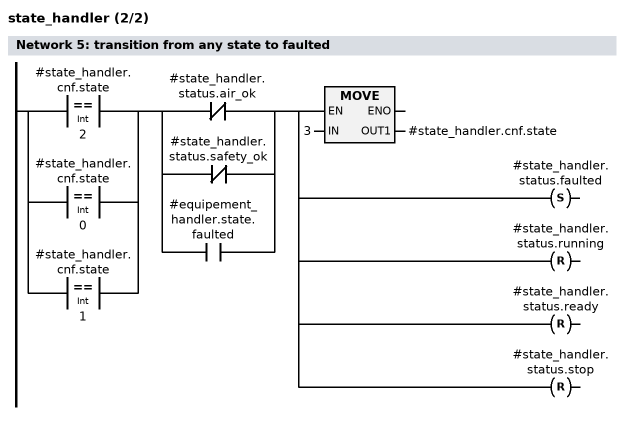
   RUNG wire#powerrail
      { S7_Templates := "SrcType := Int" } EQ_Contact(in1 := #state_handler.cnf.state, in2 := 2)
      wire#w1
      I_Contact( #state_handler.status.air_ok )
      wire#w2
      Move(in := 3, out1 => #state_handler.cnf.state)
   END_RUNG
   RUNG wire#powerrail
      { S7_Templates := "SrcType := Int" } EQ_Contact(in1 := #state_handler.cnf.state, in2 := 0)
   END_RUNG wire#w1
   RUNG wire#powerrail
      { S7_Templates := "SrcType := Int" } EQ_Contact(in1 := #state_handler.cnf.state, in2 := 1)
   END_RUNG wire#w1
   RUNG wire#w1
      I_Contact( #state_handler.status.safety_ok )
   END_RUNG wire#w2
   RUNG wire#w1
      Contact( #equipement_handler.state.faulted )
   END_RUNG wire#w2
   RUNG wire#w2
      S_Coil( #state_handler.status.faulted )
   END_RUNG
   RUNG wire#w2
      R_Coil( #state_handler.status.running )
   END_RUNG
   RUNG wire#w2
      R_Coil( #state_handler.status.ready )
   END_RUNG
   RUNG wire#w2
      R_Coil( #state_handler.status.stop )
   END_RUNG
   // the same network as SCL:
   #_w1 := ((#state_handler.cnf.state = 2) OR (#state_handler.cnf.state = 0) OR (#state_handler.cnf.state = 1)) AND (NOT #state_handler.status.air_ok OR NOT #state_handler.status.safety_ok OR #equipement_handler.state.faulted);
   IF #_w1 THEN
       #state_handler.cnf.state := 3;
       #state_handler.status.faulted := TRUE;
       #state_handler.status.running := FALSE;
       #state_handler.status.ready := FALSE;
       #state_handler.status.stop := FALSE;
   END_IF;
END_REGION
END_FUNCTION_BLOCK

FUNCTION_BLOCK "tower_handler"   // FB3, LAD
{ S7_Optimized_Access := 'TRUE' }
VERSION : 0.1
   VAR_OUTPUT
      tower_green_light : Bool;
      tower_red_light : Bool;
      tower_orange_light : Bool;
      tower_buzer : Bool;
   END_VAR
   VAR_IN_OUT
      state_handler_Machine : "udt_state_handler";
      tower_udt : "udt_tower_handler";
   END_VAR
BEGIN

REGION Network 1: geen light machine is running
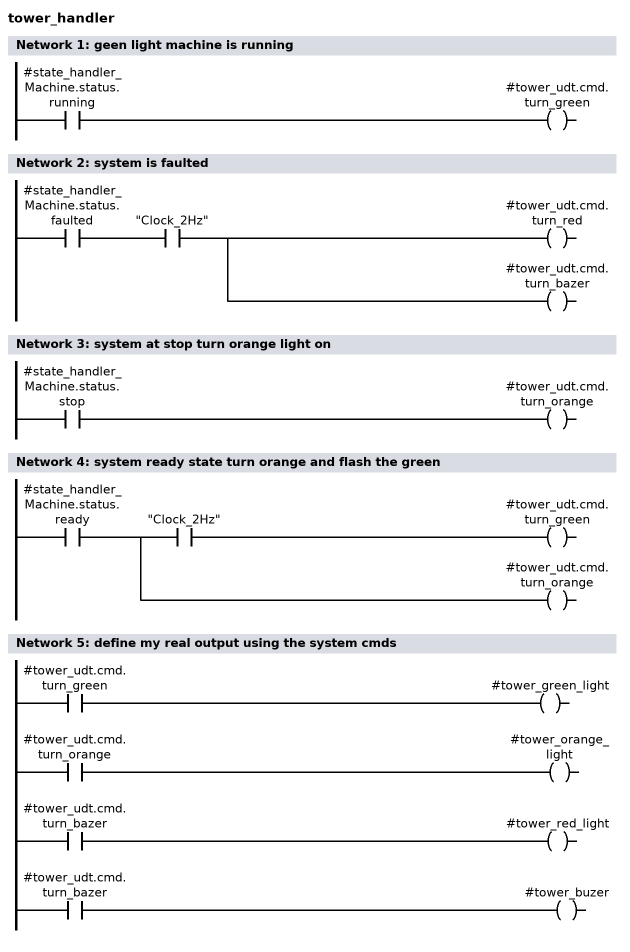
   RUNG wire#powerrail
      Contact( #state_handler_Machine.status.running )
      Coil( #tower_udt.cmd.turn_green )
   END_RUNG
   // the same network as SCL:
   #tower_udt.cmd.turn_green := #state_handler_Machine.status.running;
END_REGION

REGION Network 2: system is faulted
   RUNG wire#powerrail
      Contact( #state_handler_Machine.status.faulted )
      Contact( "Clock_2Hz" )
      wire#w1
      Coil( #tower_udt.cmd.turn_red )
   END_RUNG
   RUNG wire#w1
      Coil( #tower_udt.cmd.turn_bazer )
   END_RUNG
   // the same network as SCL:
   #tower_udt.cmd.turn_red := #state_handler_Machine.status.faulted AND "Clock_2Hz";
   #tower_udt.cmd.turn_bazer := #tower_udt.cmd.turn_red;
END_REGION

REGION Network 3: system at stop turn orange light on
   RUNG wire#powerrail
      Contact( #state_handler_Machine.status.stop )
      Coil( #tower_udt.cmd.turn_orange )
   END_RUNG
   // the same network as SCL:
   #tower_udt.cmd.turn_orange := #state_handler_Machine.status.stop;
END_REGION

REGION Network 4: system ready state turn orange and flash the green
   RUNG wire#powerrail
      Contact( #state_handler_Machine.status.ready )
      wire#w1
      Contact( "Clock_2Hz" )
      Coil( #tower_udt.cmd.turn_green )
   END_RUNG
   RUNG wire#w1
      Coil( #tower_udt.cmd.turn_orange )
   END_RUNG
   // the same network as SCL:
   #tower_udt.cmd.turn_green := #state_handler_Machine.status.ready AND "Clock_2Hz";
   #tower_udt.cmd.turn_orange := #state_handler_Machine.status.ready;
END_REGION

REGION Network 5: define my real output using the system cmds
   RUNG wire#powerrail
      Contact( #tower_udt.cmd.turn_green )
      Coil( #tower_green_light )
   END_RUNG
   RUNG wire#powerrail
      Contact( #tower_udt.cmd.turn_orange )
      Coil( #tower_orange_light )
   END_RUNG
   RUNG wire#powerrail
      Contact( #tower_udt.cmd.turn_bazer )
      Coil( #tower_red_light )
   END_RUNG
   RUNG wire#powerrail
      Contact( #tower_udt.cmd.turn_bazer )
      Coil( #tower_buzer )
   END_RUNG
   // the same network as SCL:
   #tower_green_light := #tower_udt.cmd.turn_green;
   #tower_orange_light := #tower_udt.cmd.turn_orange;
   #tower_red_light := #tower_udt.cmd.turn_bazer;
   #tower_buzer := #tower_udt.cmd.turn_bazer;
END_REGION
END_FUNCTION_BLOCK

FUNCTION_BLOCK "safety_block"   // FB4, LAD
{ S7_Optimized_Access := 'TRUE' }
VERSION : 0.1
   VAR_INPUT
      reset : Bool;
      emg_stop : Bool;
   END_VAR
   VAR_IN_OUT
      state_handler : "udt_state_handler";
   END_VAR
   VAR_TEMP
      reset_pulse_safety : Bool;
   END_VAR
   VAR_TEMP   // added for the SCL form of the ladder/FBD networks
      _w1 : Bool;
      _w2 : Bool;
   END_VAR
BEGIN

REGION Network 1: watch emergency stop
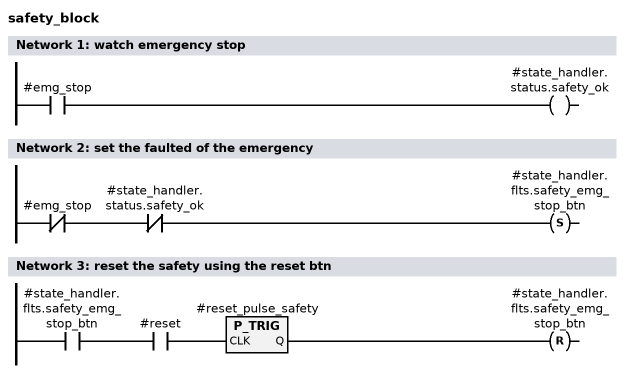
   RUNG wire#powerrail
      Contact( #emg_stop )
      Coil( #state_handler.status.safety_ok )
   END_RUNG
   // the same network as SCL:
   #state_handler.status.safety_ok := #emg_stop;
END_REGION

REGION Network 2: set the faulted of the emergency
   RUNG wire#powerrail
      I_Contact( #emg_stop )
      I_Contact( #state_handler.status.safety_ok )
      S_Coil( #state_handler.flts.safety_emg_stop_btn )
   END_RUNG
   // the same network as SCL:
   IF NOT #emg_stop AND NOT #state_handler.status.safety_ok THEN
       #state_handler.flts.safety_emg_stop_btn := TRUE;
   END_IF;
END_REGION

REGION Network 3: reset the safety using the reset btn
   RUNG wire#powerrail
      Contact( #state_handler.flts.safety_emg_stop_btn )
      Contact( #reset )
      P_Trig( #reset_pulse_safety )
      R_Coil( #state_handler.flts.safety_emg_stop_btn )
   END_RUNG
   // the same network as SCL:
   #_w1 := #state_handler.flts.safety_emg_stop_btn AND #reset;
   #_w2 := #_w1 AND NOT #reset_pulse_safety;   // rising edge
   #reset_pulse_safety := #_w1;
   IF #_w2 THEN #state_handler.flts.safety_emg_stop_btn := FALSE; END_IF;
END_REGION
END_FUNCTION_BLOCK

FUNCTION_BLOCK "air_management_blk"   // FB5, LAD
{ S7_Optimized_Access := 'TRUE' }
VERSION : 0.1
   VAR_INPUT
      reset_btn : Bool;
      air_switch : Bool;
      valve_open_fb : Bool;
   END_VAR
   VAR_OUTPUT
      main_air_valve : Bool;
   END_VAR
   VAR_IN_OUT
      state_handler : "udt_state_handler";
   END_VAR
   VAR
      state : Int;
      air_start_cmd : Bool;
      air_faulted : Bool;
   END_VAR
   VAR_TEMP
      reset_pulse : Bool;
   END_VAR
   VAR_TEMP   // added for the SCL form of the ladder/FBD networks
      _w1 : Bool;
      _w2 : Bool;
   END_VAR
BEGIN

REGION Network 1: trigger the fault if the air is not enabled when cmd is there using 1min timer
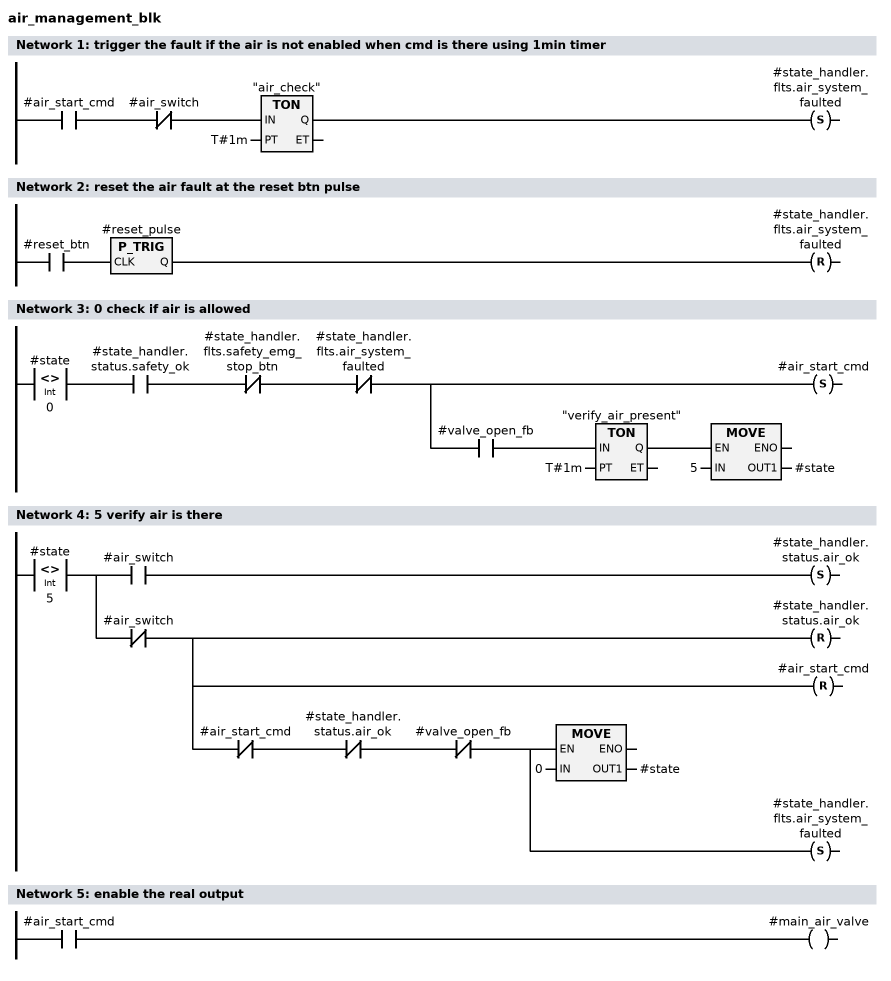
   "air_check".TON(IN := #air_start_cmd AND NOT #air_switch, PT := T#1m);
   IF "air_check".Q THEN #state_handler.flts.air_system_faulted := TRUE; END_IF;
END_REGION

REGION Network 2: reset the air fault at the reset btn pulse
   RUNG wire#powerrail
      Contact( #reset_btn )
      P_Trig( #reset_pulse )
      R_Coil( #state_handler.flts.air_system_faulted )
   END_RUNG
   // the same network as SCL:
   #_w1 := #reset_btn AND NOT #reset_pulse;   // rising edge
   #reset_pulse := #reset_btn;
   IF #_w1 THEN #state_handler.flts.air_system_faulted := FALSE; END_IF;
END_REGION

REGION Network 3: 0 check if air is allowed
   #_w1 := (#state <> 0) AND #state_handler.status.safety_ok AND NOT #state_handler.flts.safety_emg_stop_btn AND NOT #state_handler.flts.air_system_faulted;
   IF #_w1 THEN #air_start_cmd := TRUE; END_IF;
   "verify_air_present".TON(IN := #_w1 AND #valve_open_fb, PT := T#1m);
   IF "verify_air_present".Q THEN #state := 5; END_IF;
END_REGION

REGION Network 4: 5 verify air is there
   RUNG wire#powerrail
      { S7_Templates := "SrcType := Int" } NE_Contact(in1 := #state, in2 := 5)
      wire#w1
      Contact( #air_switch )
      S_Coil( #state_handler.status.air_ok )
   END_RUNG
   RUNG wire#w1
      I_Contact( #air_switch )
      wire#w2
      R_Coil( #state_handler.status.air_ok )
   END_RUNG
   RUNG wire#w2
      R_Coil( #air_start_cmd )
   END_RUNG
   RUNG wire#w2
      I_Contact( #air_start_cmd )
      I_Contact( #state_handler.status.air_ok )
      I_Contact( #valve_open_fb )
      wire#w3
      Move(in := 0, out1 => #state)
   END_RUNG
   RUNG wire#w3
      S_Coil( #state_handler.flts.air_system_faulted )
   END_RUNG
   // the same network as SCL:
   #_w1 := #state <> 5;
   IF #_w1 AND #air_switch THEN #state_handler.status.air_ok := TRUE; END_IF;
   #_w2 := #_w1 AND NOT #air_switch;
   IF #_w2 THEN
       #state_handler.status.air_ok := FALSE;
       #air_start_cmd := FALSE;
   END_IF;
   IF #_w2 AND NOT #air_start_cmd AND NOT #state_handler.status.air_ok AND NOT #valve_open_fb THEN
       #state := 0;
       #state_handler.flts.air_system_faulted := TRUE;
   END_IF;
END_REGION

REGION Network 5: enable the real output
   RUNG wire#powerrail
      Contact( #air_start_cmd )
      Coil( #main_air_valve )
   END_RUNG
   // the same network as SCL:
   #main_air_valve := #air_start_cmd;
END_REGION
END_FUNCTION_BLOCK

FUNCTION "main_block" : Void   // FC1, LAD
{ S7_Optimized_Access := 'TRUE' }
VERSION : 0.1
BEGIN

REGION Network 1: call state handler generic block
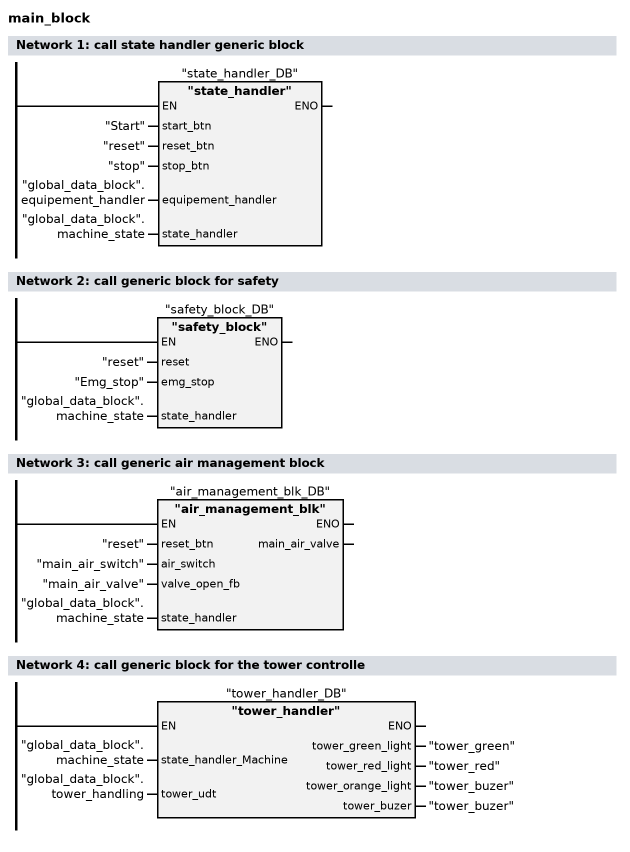
   RUNG wire#powerrail
      "state_handler_DB"(start_btn := "Start", reset_btn := "reset", stop_btn := "stop", equipement_handler := "global_data_block".equipement_handler, state_handler := "global_data_block".machine_state)
   END_RUNG
   // the same network as SCL:
   "state_handler_DB"(start_btn := "Start",   // "state_handler"
                      reset_btn := "reset",
                      stop_btn := "stop",
                      equipement_handler := "global_data_block".equipement_handler,
                      state_handler := "global_data_block".machine_state);
END_REGION

REGION Network 2: call generic block for safety
   RUNG wire#powerrail
      "safety_block_DB"(reset := "reset", emg_stop := "Emg_stop", state_handler := "global_data_block".machine_state)
   END_RUNG
   // the same network as SCL:
   "safety_block_DB"(reset := "reset",   // "safety_block"
                     emg_stop := "Emg_stop",
                     state_handler := "global_data_block".machine_state);
END_REGION

REGION Network 3: call generic air management block
   RUNG wire#powerrail
      "air_management_blk_DB"(reset_btn := "reset", air_switch := "main_air_switch", valve_open_fb := "main_air_valve", state_handler := "global_data_block".machine_state, main_air_valve =>)
   END_RUNG
   // the same network as SCL:
   "air_management_blk_DB"(reset_btn := "reset",   // "air_management_blk"
                           air_switch := "main_air_switch",
                           valve_open_fb := "main_air_valve",
                           state_handler := "global_data_block".machine_state);
END_REGION

REGION Network 4: call generic block for the tower controlle
   RUNG wire#powerrail
      "tower_handler_DB"(state_handler_Machine := "global_data_block".machine_state, tower_udt := "global_data_block".tower_handling, tower_green_light => "tower_green", tower_red_light => "tower_red", tower_orange_light => "tower_buzer", tower_buzer => "tower_buzer")
   END_RUNG
   // the same network as SCL:
   "tower_handler_DB"(state_handler_Machine := "global_data_block".machine_state,   // "tower_handler"
                      tower_udt := "global_data_block".tower_handling,
                      tower_green_light => "tower_green",
                      tower_red_light => "tower_red",
                      tower_orange_light => "tower_buzer",
                      tower_buzer => "tower_buzer");
END_REGION
END_FUNCTION

(* ===== HMI "HMI_RT_1" =====
system functions are stored by id; their names below are inferred from use
connection "HMI_Connection_1": ETHERNET, S7_1500_OMS

HMI tags "Default tag table"
   "bottle_movement" : Int, internal
   "screen_number" : Int, internal
   "box_at_filling" : Bool = PLC box_at_filling AT %I1.0, 1 s
   "box_at_sealing" : Bool = PLC part_at_sealing AT %I3.2, 1 s
   "box_at_reject" : Bool = PLC box_at_reject AT %I5.1, 1 s
   "box_had_left" : Bool = PLC box_left AT %I1.3, 1 s
   "box_rejected" : Bool = PLC box_reject AT %I1.2, 1 s
   "box_at_scale" : Bool = PLC box_at_scale AT %I1.1, 1 s
   "1_main_squence_DB_bottle_count_done" : Int = PLC "1_main_squence_DB".bottle_count_done, 1 s
   "global_data_block_verification_handler_status_pass_part" : Bool = PLC global_data_block.verification_handler.status.pass_part, 1 s
   "global_data_block_verification_handler_status_reject_part" : Bool = PLC global_data_block.verification_handler.status.reject_part, 1 s
   "global_data_block_verification_handler_status_actual_weight_bottle" : Int = PLC global_data_block.verification_handler.status.actual_weight_bottle, 1 s
   "curent_speed" : Word = PLC curent_speed AT %IW600, 1 s
   "set_point_vfd" : Word = PLC set_point_vfd AT %QW600, 1 s
   "global_data_block_hmi_cmd_state_cmd_oprator_speed_setpoint" : Int = PLC global_data_block.hmi_cmd_state.cmd.oprator_speed_setpoint, 1 s
   "global_data_block_filling_station_handler_flt1" : Word = PLC global_data_block.filling_station_handler.flt1, 1 s
   "global_data_block_filling_station_handler_flt2" : Word = PLC global_data_block.filling_station_handler.flt2, 1 s
   "global_data_block_sealing_handler_flt_locater_cylinder" : Word = PLC global_data_block.sealing_handler.flt_locater_cylinder, 1 s
   "global_data_block_sealing_handler_flt_valve_carrier_cyl" : Word = PLC global_data_block.sealing_handler.flt_valve_carrier_cyl, 1 s
   "global_data_block_filling_station_handler_flt_valve" : Word = PLC global_data_block.filling_station_handler.flt_valve, 1 s
   "global_data_block_sealing_handler_flt_valve" : Word = PLC global_data_block.sealing_handler.flt_valve, 1 s
   "global_data_block_reject_handler_flt" : Word = PLC global_data_block.reject_handler.flt, 1 s
   "safety_block_DB_emg_stop" : Bool = PLC safety_block_DB.emg_stop, 1 s

HMI tags "Tag table_1"
   "machine_running" : Bool = PLC global_data_block.machine_state.status.running AT %DB1.DBW0, 1 s
   "machine_stop" : Bool = PLC global_data_block.machine_state.status.stop AT %DB1.DBW0, 1 s
   "machine_ready" : Bool = PLC global_data_block.machine_state.status.ready AT %DB1.DBW0, 1 s
   "machine_faulted" : Bool = PLC global_data_block.machine_state.status.faulted AT %DB1.DBW0, 1 s
   "tower_cmd_green" : Bool = PLC global_data_block.tower_handling.cmd.turn_green AT %DB1.DBX0.0, 1 s
   "tower_cmd_orange" : Bool = PLC global_data_block.tower_handling.cmd.turn_orange AT %DB1.DBX0.0, 1 s
   "tower_cmd_red" : Bool = PLC global_data_block.tower_handling.cmd.turn_red AT %DB1.DBX0.0, 1 s
   "filling_cyl_extend" : Bool = PLC filling_cyl_extended AT %I4.1, 1 s
   "fillinfig_cyl_retract" : Bool = PLC filling_cyl_retracted AT %I4.0, 1 s
   "filling_carrier_valve_extended" : Bool = PLC filling_valve_extended AT %I4.4, 1 s
   "filling_carrier_valve_retracted" : Bool = PLC filling_valve_retracted AT %I4.5, 1 s
   "sealing_cyl_locater_extended" : Bool = PLC sealing_locater_extended AT %I4.6, 1 s
   "sealing_cyl_locater_retracted" : Bool = PLC sealing_locater_retacted AT %I4.7, 1 s
   "sealing_cyl_capCarrier_retracted" : Bool = PLC cap_carrier_retracted AT %I4.3, 1 s
   "sealing_capCarrier_cyl_extended" : Bool = PLC cap_carrier_extended AT %I4.2, 1 s
   "reject_cyl_retracted" : Bool = PLC reject_cyl_retracted AT %I1.5, 1 s
   "reject_cyl_extended" : Bool = PLC reject_cyl_extended AT %I1.4, 1 s
   "filling_valve" : Bool = PLC valve_switch_open AT %I2.2, 1 s
   "sealing_valve" : Bool = PLC cap_valve_open AT %I5.0, 1 s
   "conveyer_on" : Bool = PLC conveyer_moving AT %I2.1, 1 s
   "bottle_total_count" : Int = PLC "1_main_squence_DB".bottle_count_done AT %DB1.DBW0, 1 s

HMI tags "Tag table_2"
   "start_machine_cmd" : Bool = PLC global_data_block.machine_state.cmd.start AT %DB1.DBX0.0, 1 s
   "stop_cmd" : Bool = PLC global_data_block.machine_state.cmd.stop AT %DB1.DBW0, 1 s
   "reset_cmd" : Bool = PLC global_data_block.machine_state.cmd.reset AT %DB1.DBW0, 1 s

discrete alarms
   1: 'filling locater didn't reach position retracted', class Errors, trigger "global_data_block_filling_station_handler_flt1" bit 0
   2: 'filling locater didn't reach position extended', class Errors, trigger "global_data_block_filling_station_handler_flt1" bit 1
   3: 'filling valve failed to reach fillling valve failed to reachretract position', class Errors, trigger "global_data_block_filling_station_handler_flt2" bit 0
   4: 'valve filling cylinder failed to reach extended position', class Errors, trigger "global_data_block_filling_station_handler_flt2" bit 1
   5: 'cap cylinder locater failed to reach it extended position', class Errors, trigger "global_data_block_sealing_handler_flt_locater_cylinder" bit 0
   6: 'capping cyl locater failed to reach it retract position', class Errors, trigger "global_data_block_sealing_handler_flt_locater_cylinder" bit 1
   7: 'capping cyl failed to reach it extended position', class Errors, trigger "global_data_block_sealing_handler_flt_valve_carrier_cyl" bit 0
   8: 'capping cly failed to reach retract position', class Errors, trigger "global_data_block_sealing_handler_flt_valve_carrier_cyl" bit 1
   9: 'filling valve failed to open', class Errors, trigger "global_data_block_filling_station_handler_flt_valve" bit 0
   10: 'capping valve failed to open', class Errors, trigger "global_data_block_sealing_handler_flt_valve" bit 0
   11: 'reject cyl failed to reack retract position', class Errors, trigger "global_data_block_reject_handler_flt" bit 0
   12: 'reject cyl failed to reack exteneded position', class Errors, trigger "global_data_block_reject_handler_flt" bit 1

Template "Template_1" 800x420
   Button "Exit" at 709,358 size 78x58; TextOff 'Exit'; PictureOff "ExitRuntime_TP700_Comfort_TR"; PictureOn "ExitRuntime_TP700_Comfort_TR"
      on Release: StopRuntime(0)
      on Click: function_be740847(30)
   Button "Template_Button_1" at 709,88 size 78x58; TextOff 'Auto/Man'
   Button "Template_Button_2" at 709,155 size 78x58; TextOff 'Start'
      Appearance <- "start_machine_cmd"
      on Press: SetBit("start_machine_cmd")
      on Release: ResetBit("start_machine_cmd")
   Button "Template_Button_3" at 709,223 size 78x58; TextOff 'stop'
      Appearance <- "stop_cmd"
      on Press: SetBit("stop_cmd")
      on Release: ResetBit("stop_cmd")
   Button "Template_Button_4" at 709,288 size 78x58; TextOff 'Reset'
      on Press: SetBit("reset_cmd")
      on Release: ResetBit("reset_cmd")
   Button "Template_Button_5" at 370,355 size 78x58; TextOff 'sealing'
      on Click: ActivateScreen("sealing", 4)
   Button "Template_Button_6" at 245,355 size 78x58; TextOff 'filling'
      on Click: ActivateScreen("filling", 3)
   Button "Template_Button_7" at 133,354 size 78x58; TextOff 'Alarm'
      on Click: ActivateScreen("alarm", 2)
   Button "Start screen" at 26,355 size 78x58; TextOff 'Start screen'; PictureOff "NavigateHome_TP700_Comfort_TR"; PictureOn "NavigateHome_TP700_Comfort_TR"
      on Release: ActivateScreen("home", 0)
      on Click: ActivateScreen("home", 1)
   Ellipse "Template_Ellipse_1" at 487,353 size 12x14
      Appearance <- "machine_running"
   Ellipse "Template_Ellipse_2" at 487,377 size 12x14
      Appearance <- "machine_stop"
   Ellipse "Template_Ellipse_3" at 487,401 size 12x14
      Appearance <- "machine_ready"
   Ellipse "Template_Ellipse_4" at 602,353 size 12x14
      Appearance <- "machine_faulted"
   TextField "Template_Text field_1" at 508,345 size 97x30; Text 'Running'
   TextField "Template_Text field_2" at 508,368 size 89x29; Text 'Stopped'
   TextField "Template_Text field_3" at 508,393 size 96x25; Text 'Ready'
   TextField "Template_Text field_4" at 617,344 size 86x29; Text 'Faulted'
   Rectangle "Template_Rectangle_6" at 736,7 size 25x14
      Appearance <- "tower_cmd_green"
   Rectangle "Template_Rectangle_7" at 736,22 size 25x20
      Appearance <- "tower_cmd_red"
   Rectangle "Template_Rectangle_8" at 736,40 size 25x16
      Appearance <- "tower_cmd_orange"

screen "home" 800x420, template "Template_1"
   SymbolLibrary "Symbol library_2" at 13,224 size 35x66
   SymbolLibrary "Symbol library_1" at 16,198 size 680x36
   Ellipse "Ellipse_1" at 56,262 size 16x16
      Appearance <- "conveyer_on"
   TextField "Text field_1" at 0,295 size 114x25; Text 'Main Conveyer'
   SymbolLibrary "Symbol library_4" at 72,81 size 17x25
   SymbolLibrary "Symbol library_5" at 88,93 size 79x13
   SymbolLibrary "Symbol library_6" at 166,93 size 23x25
   SymbolLibrary "Symbol library_3" at 29,10 size 97x79
   Bar "Bar_1" at 31,15 size 93x46; MinimumValue 0; MaximumValue 100
   SymbolLibrary "Symbol library_7" at 586,257 size 110x77
   TextField "Text field_2" at 72,116 size 105x17; Text 'Filling valve'
   TextField "Text field_3" at 128,27 size 102x23; Text 'reservoir'
   Circle "Circle_1" at 140,138 size 9x9
      Appearance <- "filling_valve"
   SymbolLibrary "Symbol library_8" at 147,159 size 19x28
   SymbolLibrary "Symbol library_9" at 282,158 size 19x28
   SymbolLibrary "Symbol library_10" at 404,159 size 19x28
   SymbolLibrary "Symbol library_11" at 496,159 size 19x28
   SymbolLibrary "Symbol library_12" at 606,159 size 19x28
   SymbolLibrary "Symbol library_13" at 114,187 size 19x29
      HorizontalMovement <- "bottle_movement"
   Circle "Circle_2" at 166,174 size 11x11
      Appearance <- "box_at_filling"
   Circle "Circle_3" at 301,177 size 11x11
      Appearance <- "box_at_sealing"
   Circle "Circle_4" at 422,176 size 11x11
      Appearance <- "box_at_scale"
   Circle "Circle_5" at 517,175 size 11x11
      Appearance <- "box_at_reject"
   Circle "Circle_6" at 625,174 size 11x11
      Appearance <- "box_had_left"
   SymbolLibrary "Symbol library_14" at 155,136 size 36x20
   SymbolLibrary "Symbol library_16" at 277,69 size 35x59
   SymbolLibrary "Symbol library_15" at 268,50 size 36x20
   Circle "Circle_7" at 343,83 size 14x14
      Appearance <- "sealing_cyl_capCarrier_retracted"
   Circle "Circle_8" at 343,176 size 14x14
      Appearance <- "sealing_capCarrier_cyl_extended"
   TextField "Text field_4" at 356,82 size 54x15; Text 'retract'
   TextField "Text field_5" at 356,174 size 57x15; Text 'extend'
   TextField "Text field_6" at 247,111 size 58x17; Text 'cap_M'
   SymbolLibrary "Symbol library_17" at 177,117 size 13x21
   TextField "Text field_7" at 387,199 size 68x17; Text 'scale'
   IOField "I/O field_1" at 365,239 size 89x31; FormatPattern s9999; Unit  g
      ProcessValue <- "global_data_block_verification_handler_status_actual_weight_bottle"
   TextField "Text field_8" at 365,285 size 87x14; Text 'part_passed'
   TextField "Text field_9" at 365,311 size 90x21; Text 'part_rejected'
   Circle "Circle_9" at 454,288 size 9x9
      Appearance <- "global_data_block_verification_handler_status_pass_part"
   Circle "Circle_10" at 453,315 size 9x9
      Appearance <- "global_data_block_verification_handler_status_reject_part"
   SymbolLibrary "Symbol library_18" at 178,149 size 13x21
   TextField "Text field_10" at 301,32 size 82x28; Text 'cap_valve'
   Circle "Circle_11" at 508,59 size 9x9
      Appearance <- "reject_cyl_retracted"
   Circle "Circle_12" at 508,124 size 9x9
      Appearance <- "reject_cyl_extended"
   TextField "Text field_11" at 518,56 size 58x19; Text 'retract'
   TextField "Text field_12" at 518,121 size 59x20; Text 'extend'
   TextField "Text field_13" at 460,19 size 110x26; Text 'reject_cylinder'
   TextField "Text field_14" at 578,52 size 115x31; Text 'Bottle count'
   IOField "I/O field_3" at 598,106 size 75x31; FormatPattern s9999
      ProcessValue <- "1_main_squence_DB_bottle_count_done"
   Circle "Circle_13" at 215,137 size 14x14
      Appearance <- "filling_carrier_valve_retracted"
   Circle "Circle_14" at 215,175 size 14x14
      Appearance <- "filling_carrier_valve_extended"
   Circle "Circle_15" at 252,57 size 14x14
      Appearance <- "sealing_valve"
   TextField "Text field_15" at 190,238 size 136x23; Text 'VFD Data'
   IOField "I/O field_2" at 214,265 size 115x31; FormatPattern 99999; Unit  rpm
      ProcessValue <- "curent_speed"
   IOField "I/O field_4" at 215,298 size 113x31; FormatPattern s99999; Unit  %
      ProcessValue <- "global_data_block_hmi_cmd_state_cmd_oprator_speed_setpoint"
   TextField "Text field_16" at 116,271 size 102x29; Text 'Actual speed'
   TextField "Text field_17" at 115,299 size 99x26; Text 'Set point s'

screen "alarm" 800x420, template "Template_1"
   AlarmView "Alarm view_1" at 1,7 size 692x334

VB script "VBFunction_1"
   'Tip:
   ' 1. Use the <CTRL+SPACE> or <CTRL+I> shortcut to open a list of all objects and functions
   ' 2. Write the code using the HMI Runtime object.
   '  Example: HmiRuntime.Screens("Screen_1").
   ' 3. Use the <CTRL+J> shortcut to create an object reference.
   'Write the code as of this position:
*)